// TIA Portal V20 export
// export: Created 2026-10-11T05:22:25.6370833Z, ExportSetting WithDefaults, DisplayName Totally Integrated Automation Portal, DisplayVersion V20, DisplayName TIA Portal Openness, DisplayVersion V20, DisplayName TIA Portal Teamcenter Gateway, DisplayVersion V20, DisplayName TIA Portal Version Control Interface, DisplayVersion V20, DisplayName SINAMICS Startdrive Advanced, DisplayVersion V20 SP1 Update 2, DisplayName SINAMICS Startdrive G110M, G120, G120C, G120D, G120P, G115D, DisplayVersion V20 SP1 Update 2, DisplayName SINAMICS Startdrive G130, G150, S120, S150, SINAMICS MV, G220, S200, S210, DisplayVersion V20 SP1 Update 2, DisplayName STEP 7 Professional, DisplayVersion V20, DisplayName STEP 7 Safety, DisplayVersion V20, DisplayName WinCC Basic/Comfort/Advanced, DisplayVersion V20, DisplayName WinCC Professional, DisplayVersion V20, DisplayName WinCC Unified, DisplayVersion V20
FUNCTION "FRK_ReleaseReason" : Void   // FC42, SCL
{ S7_Optimized_Access := 'TRUE' }
VERSION : 0.1
// stored: AutoNumber true, IsIECCheckEnabled false, SetENOAutomatically false, UDAEnableTagReadback false
   VAR_INPUT
      Description : WString;
      Reason : DInt;
      Path : WString;
      Kind : DInt;
   END_VAR
   VAR_IN_OUT
      Report : "ST_ReleaseReport";
   END_VAR
BEGIN

   #Report.Released := FALSE;
   IF #Report.Count < 24 THEN
       #Report.Count := #Report.Count + 1;
       #Report.Reasons[#Report.Count].Description := #Description;
       #Report.Reasons[#Report.Count].ReasonCode := #Reason;
       #Report.Reasons[#Report.Count].SourcePath := #Path;
       #Report.Reasons[#Report.Count].Kind := #Kind;
       #Report.Reasons[#Report.Count].Bypassable := FALSE;
   END_IF;
END_FUNCTION
